// TwinCAT 3 PLC project StorageControl
// ProgramVersion: 3.1.4026.27
// libraries:
//   Tc2_Standard, * (Beckhoff Automation GmbH)
//   Tc2_System, * (Beckhoff Automation GmbH)
// project tree:
//   / PlcTask.TcTTO
//   POUs/ MAIN.TcPOU
// real-time tasks:
//   TASK PlcTask: cycle T#10ms, priority 20, ADS port 350
// I/O:
//   DEVICE Device 1 (EtherCAT), AmsNetId 10.180.10.242.2.1

CONFIGURATION StorageControl
    RESOURCE PLC ON TwinCAT3
        TASK PlcTask(INTERVAL := T#10ms, PRIORITY := 20);
        PROGRAM MAIN WITH PlcTask : MAIN;
    END_RESOURCE
END_CONFIGURATION

// ---- POUs/MAIN.TcPOU
PROGRAM MAIN
VAR
    B1        AT %I* : BOOL;  // Nr. 5,  B1: reference switch horizontal axis
    B2         AT %I* : BOOL;  // Nr. 6,  B2: light-barrier inside
    B3        AT %I* : BOOL;  // Nr. 7,  B3: light-barrier outside
    B4          AT %I* : BOOL;  // Nr. 8,  B4: reference switch vertical axis
    B5        AT %I* : BOOL;  // Nr. 11, B5: encoder horizontal axis impulse 1
    B6        AT %I* : BOOL;  // Nr. 12, B6: encoder horizontal axis impulse 2
    B7          AT %I* : BOOL;  // Nr. 13, B7: encoder vertical axis impulse 1
    B8          AT %I* : BOOL;  // Nr. 14, B8: encoder vertical axis impulse 2
    B9   AT %I* : BOOL;  // Nr. 15, B9: reference switch cantilever front
    B10    AT %I* : BOOL;  // Nr. 16, B10: reference switch cantilever back
 
    // ---------------- OUTPUTS ----------------
    M1_Forward            AT %Q* : BOOL;  // Nr. 17, Q1 (M1): motor conveyor belt forward
    M1_Back           AT %Q* : BOOL;  // Nr. 18, Q2 (M1): motor conveyor belt backward
    M2_Forward           AT %Q* : BOOL;  // Nr. 19, Q3 (M2): motor horizontal towards rack
    M2_Back       AT %Q* : BOOL;  // Nr. 20, Q4 (M2): motor horizontal towards conveyor belt
    M3_Down               AT %Q* : BOOL;  // Nr. 21, Q5 (M3): motor vertical axis downward
    M3_Up                 AT %Q* : BOOL;  // Nr. 22, Q6 (M3): motor vertical axis upward
    M4_Forward          AT %Q* : BOOL;  // Nr. 23, Q7 (M4): motor cantilever forward
    M4_Back         AT %Q* : BOOL;  // Nr. 24, Q8 (M4): motor cantilever backward
END_VAR

ACTION Storage_Main:
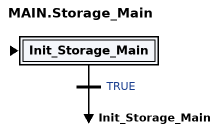
INITIAL_STEP Init_Storage_Main:
END_STEP
TRANSITION FROM Init_Storage_Main TO Init_Storage_Main
    := TRUE;
END_TRANSITION
END_ACTION

END_PROGRAM
